// TIA Portal V21 export
// export: Created 2026-11-10T07:35:23.0867044Z, ExportSetting WithDefaults, DisplayName Totally Integrated Automation Portal, DisplayVersion V21 Update 3, DisplayName STEP 7 Professional, DisplayVersion V21 Update 3, DisplayName STEP 7 Safety, DisplayVersion V21, DisplayName Tech WebApplication, DisplayVersion V21, DisplayName WinCC Basic/Comfort/Advanced, DisplayVersion V21 Update 3, DisplayName WinCC Unified, DisplayVersion V21 Update 3
FUNCTION_BLOCK "FB_Lad_ex154"   // FB56, LAD
{ S7_Optimized_Access := 'TRUE' }
VERSION : 0.1
// stored: AutoNumber true, IsIECCheckEnabled false, IsRetainMemResEnabled false, MemoryReserve 100, SetENOAutomatically false, UDAEnableTagReadback false
   VAR_INPUT
      v_ioid : Byte;
      v_addr : Word;
      v_ret_val : Int;
   END_VAR
   VAR_OUTPUT
      v_hwid : HW_IO;
   END_VAR
BEGIN

REGION Network 1: LOG2MOD - Determine the hardware identifier from addressing of STEP 7 V5.5 SPx
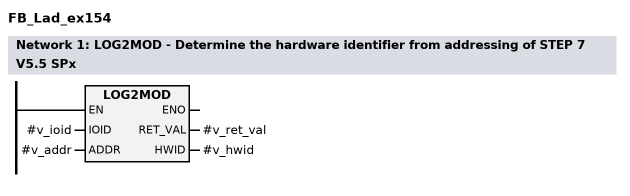
   RUNG wire#powerrail
      LOG2MOD(IOID := #v_ioid, ADDR := #v_addr, Ret_Val => #v_ret_val, HWID => #v_hwid)
   END_RUNG
   // the same network as SCL:
   #v_ret_val := LOG2MOD(IOID := #v_ioid, ADDR := #v_addr, HWID => #v_hwid);
END_REGION
END_FUNCTION_BLOCK
